FUNCTION_BLOCK FB_Fill EXTENDS FB_Base
VAR_INPUT
	bEnable   : BOOL;
	stRecipe  : ST_Recipe;
END_VAR
VAR_OUTPUT
	bDone     : BOOL;
	bError    : BOOL;
END_VAR
VAR
	fbValve   : FB_Valve;         (* bulk valve *)
	fbFine    : FB_Valve;         (* fine valve *)
	eState    : E_FillState;
	tSettle   : TIME := T#500MS;
	arrWeights : ARRAY[0..9] OF LREAL;
END_VAR

CASE eState OF
	E_FillState.Idle:
		IF bEnable THEN eState := E_FillState.Bulk; END_IF
	E_FillState.Bulk:
		fbValve.Open();
END_CASE

METHOD Start : BOOL
VAR_INPUT
	rTarget : LREAL;
END_VAR
eState := E_FillState.Bulk;
Start := TRUE;
END_METHOD

END_FUNCTION_BLOCK

(* stored: Version 1.1.0.1, ProductVersion 3.1.4024.12
   POU FB_Fill: Id {aaaaaaaa-0000-0000-0000-000000000002}, SpecialFunc None
   Method Start: Id {aaaaaaaa-0000-0000-0000-000000000003} *)
